FUNCTION F_CheckSyntaxReal : BOOL (* TRUE if STR does not contain capital letters *)
VAR_INPUT
	str 		:T_MaxString;
	flag 		:T_MaxString;
	sep 		:T_MaxString := '=';
	rsufix		:POINTER TO REAL; 					
END_VAR
VAR
	L			:INT;
	prefix1		:T_MaxString;
	prefix2		:T_MaxString;
	ssufix		:T_MaxString;
END_VAR


prefix1 := CONCAT(flag, sep);
L := LEN(prefix1);
prefix2 := MID(str, L, 1);

F_CheckSyntaxReal := FALSE;

IF LEN(str) > L
THEN
	ssufix := DELETE(str, L, 1);
	IF prefix1 = prefix2
	THEN
		IF F_CheckStringIsReal(ssufix)
		THEN
			F_CheckSyntaxReal := TRUE; 
			rsufix^ := STRING_TO_REAL(ssufix);
		END_IF
	END_IF;
END_IF

END_FUNCTION

(* stored: Version 1.1.0.1, ProductVersion 3.1.4024.15
   POU F_CheckSyntaxReal: Id {a3247213-3d66-4b3b-b3c3-a47e2f65b5b7}, SpecialFunc None *)
